Staubli VAL3: main.pgx

program main()
begin
  close(tCurrentTool)
  pPointRs.config.shoulder = lefty
  pPointRs2.config.shoulder = lefty
  mCurrentSpeed.tvel = 100.00
  mCurrentSpeed.blend = joint
  mCurrentSpeed.reach = 0.010
  mCurrentSpeed.leave = 0.010
  // Program MainCall start
  // Program generated by RoboDK v6.0.7 for Staubli TS20 FL 100 TC on XX/XX/XXXX 18:00:00
  // Using nominal kinematics.
  call MoveJoint(10.00000,-20.00000,50.00000,30.00000)
  //call prog:SubProg2()
  //call prog:NotAProgram()

  waitEndMove()
  // Program MainCall end
  // Program SubProg2 start
  call MoveJoint(30.00000,25.00000,80.00000,-45.00000)

  waitEndMove()
  // Program SubProg2 end

end
